FUNCTION_BLOCK FB_Base IMPLEMENTS ITF_Base
VAR_INPUT
END_VAR
VAR_OUTPUT
END_VAR
VAR
	nErrorId     : UDINT := 0;
    nRegisterPos : UDINT := 0;
END_VAR

{warning 'Eigenschaftenimplementierung hinzufügen'}
PROPERTY Error : UDINT
GET
Error := nErrorId;
END_GET
SET
nErrorId := Error;
END_SET
END_PROPERTY

METHOD FB_init : BOOL
VAR_INPUT
	bInitRetains : BOOL; // if TRUE, the retain variables are initialized (warm start / cold start)
	bInCopyCode : BOOL;  // if TRUE, the instance afterwards gets moved into the copy code (online change)
END_VAR
nRegisterPos := GVL.Register.AddInterfacePointer(
    ipBase := THIS^
);

FB_init := TRUE;
END_METHOD

END_FUNCTION_BLOCK

(* stored: Version 1.1.0.1, ProductVersion 3.1.4024.16
   POU FB_Base: Id {bfd93158-86fb-49c5-a29a-90f08bc218ef}, SpecialFunc None
   Property Error: Id {26298a54-29d6-43b2-959a-bbce0a92d7be}
   Get Get: Id {2fb8a451-d62c-4022-bb29-225339fca2fe}
   Set Set: Id {6d1a74c1-1abe-4f41-994c-e15f837cd29b}
   Method FB_init: Id {e19e7be8-b78a-4094-82fc-43404e66254d} *)
